(*
SPDX-FileCopyrightText: c 2026 Oleksandr Tiutyk <trofimich@gmail.com>
SPDX-License-Identifier: MIT
License: https://opensource.org/license/mit
*)

(*!
<summary>Checks copy isolation and the lifetime of a borrowed entry.</summary>
<description>
Borrows a group-owned stack reserved for this case. Use from one task at a stable address.
Teardown clears the stack and test-owned resources before publication.
</description>
*)

{attribute 'no_assign'}
{attribute 'no_explicit_call' := 'do not call this function block directly'}
FUNCTION_BLOCK StackCopiedAndBorrowedValuesTest EXTENDS TOF_Testing.SingleCycleTest
VAR_STAT
	{attribute 'hide'}
	_ClassName : STRING := __POUNAME();
END_VAR
VAR
	_Stack : TOF_Collections.IStack;
	_SourceValue : INT;
END_VAR

(*!
<summary>Clears the fixture before the runner publishes the result.</summary>
<description>
Also runs after an unexpected exception interrupts the case.
</description>
*)
METHOD PROTECTED AfterTest
_Stack.Clear();
END_METHOD

//! <summary>Borrows the concrete class name. Callers must not modify it.</summary>
{attribute 'monitoring' := 'call'}
PROPERTY ClassName : REFERENCE TO STRING
GET
ClassName REF= _ClassName;
END_GET
END_PROPERTY

(*!
<summary>Checks copy isolation and the lifetime of a borrowed entry.</summary>
*)
METHOD PROTECTED ExecuteTest
VAR
	query : TOF_Core.GENERIC_VALUE;
END_VAR
_SourceValue := 7;
_Stack.PushCopy(value := _SourceValue);
_SourceValue := 9;

Assert.ThatInt(
	actual := _Stack.Peek().AsInt(),
	message := "PushCopy must isolate the value from later source writes"
).ToBe(expected := INT#7);

query := TOF_Core.GenericValueFactory.FromIntReference(value := _SourceValue);
_Stack.PushGeneric(value := query);
_SourceValue := 11;

Assert.ThatInt(
	actual := _Stack.Peek().AsInt(),
	message := "PushGeneric must observe the current value in borrowed storage"
).ToBe(expected := INT#11);

Assert.ThatBool(
	actual := NOT _Stack.Peek().IsMemoryOwner AND_THEN _Stack.Peek().Address = query.Address,
	message := "The stored descriptor must retain the borrowed address and ownership mode"
).IsTrue();

Assert.ThatBool(
	actual := _Stack.ContainsGeneric(value := query, releaseValue := FALSE),
	message := "Borrowed lookup must find the top"
).IsTrue();

_Stack.RemoveLast();

Assert.ThatInt(
	actual := _SourceValue,
	message := "Removing a borrowed entry must preserve its source"
).ToBe(expected := INT#11);

Assert.ThatInt(
	actual := _Stack.Peek().AsInt(),
	message := "Removing the borrowed entry must reveal the copy"
).ToBe(expected := INT#7);
END_METHOD

(*!
<summary>Binds the stack fixture for this case.</summary>
<description>
Stores a borrowed interface without invoking the fixture. The owning group keeps it alive and
reserves it for this case. TestElement initializes the name and parent.
</description>
<param name="name">Display name of this case.</param>
<param name="parent">Group that owns this case.</param>
<param name="stack">Required live stack reserved for this case.</param>
*)
METHOD FB_init : BOOL
VAR_INPUT
	bInitRetains: BOOL; // TRUE: the retain variables are initialized (reset warm / reset cold)
	bInCopyCode: BOOL; // TRUE: the instance will be copied to the copy code afterward (online change)
	name : WSTRING;
	parent : TOF_Testing.ITestElement;
	stack : TOF_Collections.IStack;
END_VAR
_Stack := stack;
FB_init := TRUE;
END_METHOD

//! <summary>Borrows the compiler-initialized namespace name. Callers must not modify it.</summary>
{attribute 'monitoring' := 'call'}
PROPERTY NamespaceName : REFERENCE TO STRING
GET
NamespaceName REF= CurrentNamespace.Name;
END_GET
END_PROPERTY

//! <summary>Reports the concrete instance size in bytes.</summary>
{attribute 'monitoring' := 'call'}
PROPERTY SelfSize : ULINT
GET
SelfSize := XSIZEOF(THIS^);
END_GET
END_PROPERTY

END_FUNCTION_BLOCK

(* stored: Version 1.1.0.1, ProductVersion 3.1.4026.21
   POU StackCopiedAndBorrowedValuesTest: Id {7a6a2524-575f-4e68-8748-0298ca0c0fc2}, SpecialFunc None
   Method AfterTest: Id {039205af-7a1b-4030-87cb-f2628bbedcf3}
   Property ClassName: Id {e77cca29-49af-47ff-9072-95e58eea69c4}
   Get Get: Id {bcb4e491-9869-4c5b-a228-c129637c378d}
   Method ExecuteTest: Id {ca86fe69-ac16-4dc2-a691-db5ee98a42fc}
   Method FB_init: Id {e155ef1c-a70b-4f64-8013-3c63e03703ee}
   Property NamespaceName: Id {97da9e1f-fbb5-4291-b493-9847cfc279f4}
   Get Get: Id {235c04e5-c08f-4551-904f-a8c02deda7de}
   Property SelfSize: Id {05173312-1609-4c3f-8d5e-35c75bd144c8}
   Get Get: Id {071bdc44-b875-433a-9a02-f52914d81efd} *)
